Staubli VAL3: getSize.pgx

public program getSize(num& x_nSize, num& x_nSize1)
begin
  if io:nMaxdigital%16!=0 and nPageIndex==nPage-1
    x_nSize=io:nMaxdigital%16
  else
    x_nSize=16
  endIf
 if io:nMaxAnalog%16!=0 and nPageIndex==nPage-1
    x_nSize1=io:nMaxAnalog%16
  else
    x_nSize1=16
  endIf
end
